Fanuc TP program (LS listing): POLIR.LS

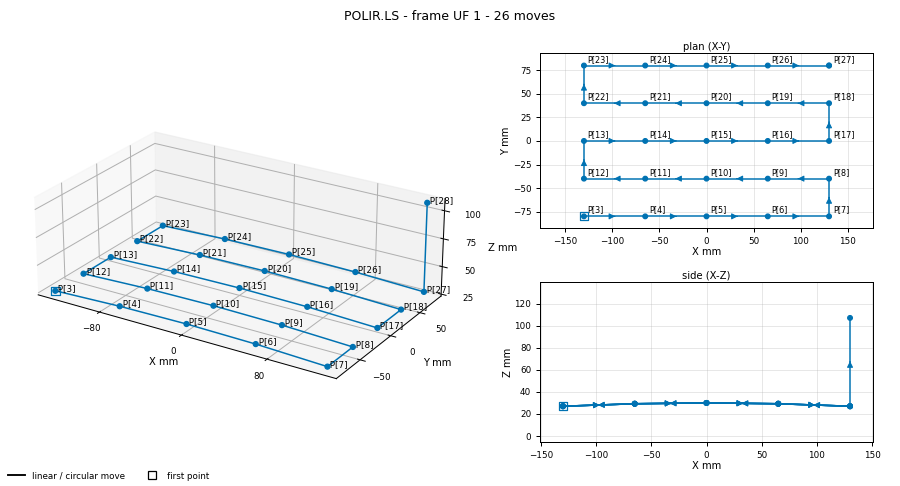
[picture p0: tool path of POLIR.LS in frame UF 1, 26 of 29 moves have a stored position in this frame; points joined in program order, loops and branches not executed]
/PROG  POLIR
/ATTR
OWNER		= MNEDITOR;
COMMENT		= "RoboDK sequence";
PROG_SIZE	= 0;
CREATE		= DATE 31-12-14  TIME 12:00:00;
MODIFIED	= DATE 31-12-14  TIME 12:00:00;
FILE_NAME	= POLIR;
VERSION		= 0;
LINE_COUNT	= 38;
MEMORY_SIZE	= 0;
PROTECT		= READ_WRITE;
TCD:  STACK_SIZE	= 0,
      TASK_PRIORITY	= 50,
      TIME_SLICE	= 0,
      BUSY_LAMP_OFF	= 0,
      ABORT_REQUEST	= 0,
      PAUSE_REQUEST	= 0;
DEFAULT_GROUP	= 1,*,*,*,*,*,*;
CONTROL_CODE	= 00000000 00000000;
/MN
   1:  ! Program generated by RoboDK v6.0.6 for FANUC M-10iD/12 on 24/ ;
   2:  ! 09/2026 00:37:20 ;
   3:  ! Using nominal kinematics. ;
   4:  UFRAME_NUM=1 ;
   5:  ! UF1:850.0,0.0,90.0,0.0,0.0,0.0 ;
   6:  UTOOL_NUM=1 ;
   7:  ! UT1:0.0,0.0,200.0,0.0,0.0,0.0 ;
   8:J P[1] 2% CNT1 ACC100 ;
   9:J P[2] 2% CNT1 ACC100 ;
  10:  DO[1]=ON ;
  11:L P[3] 40mm/sec CNT1 ACC100 ;
  12:L P[4] 40mm/sec CNT1 ACC100 ;
  13:L P[5] 40mm/sec CNT1 ACC100 ;
  14:L P[6] 40mm/sec CNT1 ACC100 ;
  15:L P[7] 40mm/sec CNT1 ACC100 ;
  16:L P[8] 40mm/sec CNT1 ACC100 ;
  17:L P[9] 40mm/sec CNT1 ACC100 ;
  18:L P[10] 40mm/sec CNT1 ACC100 ;
  19:L P[11] 40mm/sec CNT1 ACC100 ;
  20:L P[12] 40mm/sec CNT1 ACC100 ;
  21:L P[13] 40mm/sec CNT1 ACC100 ;
  22:L P[14] 40mm/sec CNT1 ACC100 ;
  23:L P[15] 40mm/sec CNT1 ACC100 ;
  24:L P[16] 40mm/sec CNT1 ACC100 ;
  25:L P[17] 40mm/sec CNT1 ACC100 ;
  26:L P[18] 40mm/sec CNT1 ACC100 ;
  27:L P[19] 40mm/sec CNT1 ACC100 ;
  28:L P[20] 40mm/sec CNT1 ACC100 ;
  29:L P[21] 40mm/sec CNT1 ACC100 ;
  30:L P[22] 40mm/sec CNT1 ACC100 ;
  31:L P[23] 40mm/sec CNT1 ACC100 ;
  32:L P[24] 40mm/sec CNT1 ACC100 ;
  33:L P[25] 40mm/sec CNT1 ACC100 ;
  34:L P[26] 40mm/sec CNT1 ACC100 ;
  35:L P[27] 40mm/sec CNT1 ACC100 ;
  36:L P[28] 40mm/sec CNT1 ACC100 ;
  37:  DO[1]=OFF ;
  38:J P[29] 2% CNT1 ACC100 ;
/POS
P[1]{
   GP1:
    UF : 1, UT : 1,
	J1=    -6.453 deg,	J2=    -8.040 deg,	J3=    -17.302 deg,
	J4=    -0.316 deg,	J5=    -70.069 deg,	J6=    6.554 deg
};
P[2]{
   GP1:
    UF : 1, UT : 1,
	J1=    -6.453 deg,	J2=    -6.370 deg,	J3=    -28.638 deg,
	J4=    -0.348 deg,	J5=    -58.733 deg,	J6=    6.627 deg
};
P[3]{
   GP1:
    UF : 1, UT : 1,        CONFIG : 'N U T, 0, 0, 0',
	X =  -130.000  mm,	Y =   -80.000  mm,	Z =    26.996  mm,
	W =   180.000 deg,	P =    -2.646 deg,	R =     0.000 deg
};
P[4]{
   GP1:
    UF : 1, UT : 1,        CONFIG : 'N U T, 0, 0, 0',
	X =   -65.000  mm,	Y =   -80.000  mm,	Z =    29.249  mm,
	W =   180.000 deg,	P =    -1.324 deg,	R =     0.000 deg
};
P[5]{
   GP1:
    UF : 1, UT : 1,        CONFIG : 'N U T, 0, 0, 0',
	X =     0.000  mm,	Y =   -80.000  mm,	Z =    30.000  mm,
	W =   180.000 deg,	P =     0.000 deg,	R =     0.000 deg
};
P[6]{
   GP1:
    UF : 1, UT : 1,        CONFIG : 'N U T, 0, 0, 0',
	X =    65.000  mm,	Y =   -80.000  mm,	Z =    29.249  mm,
	W =   180.000 deg,	P =     1.324 deg,	R =     0.000 deg
};
P[7]{
   GP1:
    UF : 1, UT : 1,        CONFIG : 'N U T, 0, 0, 0',
	X =   130.000  mm,	Y =   -80.000  mm,	Z =    26.996  mm,
	W =   180.000 deg,	P =     2.646 deg,	R =     0.000 deg
};
P[8]{
   GP1:
    UF : 1, UT : 1,        CONFIG : 'N U T, 0, 0, 0',
	X =   130.000  mm,	Y =   -40.000  mm,	Z =    26.996  mm,
	W =   180.000 deg,	P =     2.646 deg,	R =     0.000 deg
};
P[9]{
   GP1:
    UF : 1, UT : 1,        CONFIG : 'N U T, 0, 0, 0',
	X =    65.000  mm,	Y =   -40.000  mm,	Z =    29.249  mm,
	W =   180.000 deg,	P =     1.324 deg,	R =     0.000 deg
};
P[10]{
   GP1:
    UF : 1, UT : 1,        CONFIG : 'N U T, 0, 0, 0',
	X =     0.000  mm,	Y =   -40.000  mm,	Z =    30.000  mm,
	W =   180.000 deg,	P =     0.000 deg,	R =     0.000 deg
};
P[11]{
   GP1:
    UF : 1, UT : 1,        CONFIG : 'N U T, 0, 0, 0',
	X =   -65.000  mm,	Y =   -40.000  mm,	Z =    29.249  mm,
	W =   180.000 deg,	P =    -1.324 deg,	R =     0.000 deg
};
P[12]{
   GP1:
    UF : 1, UT : 1,        CONFIG : 'N U T, 0, 0, 0',
	X =  -130.000  mm,	Y =   -40.000  mm,	Z =    26.996  mm,
	W =   180.000 deg,	P =    -2.646 deg,	R =     0.000 deg
};
P[13]{
   GP1:
    UF : 1, UT : 1,        CONFIG : 'N U T, 0, 0, 0',
	X =  -130.000  mm,	Y =     0.000  mm,	Z =    26.996  mm,
	W =   180.000 deg,	P =    -2.646 deg,	R =     0.000 deg
};
P[14]{
   GP1:
    UF : 1, UT : 1,        CONFIG : 'N U T, 0, 0, 0',
	X =   -65.000  mm,	Y =     0.000  mm,	Z =    29.249  mm,
	W =   180.000 deg,	P =    -1.324 deg,	R =     0.000 deg
};
P[15]{
   GP1:
    UF : 1, UT : 1,        CONFIG : 'N U T, 0, 0, 0',
	X =     0.000  mm,	Y =     0.000  mm,	Z =    30.000  mm,
	W =   180.000 deg,	P =     0.000 deg,	R =     0.000 deg
};
P[16]{
   GP1:
    UF : 1, UT : 1,        CONFIG : 'N U T, 0, 0, 0',
	X =    65.000  mm,	Y =     0.000  mm,	Z =    29.249  mm,
	W =   180.000 deg,	P =     1.324 deg,	R =     0.000 deg
};
P[17]{
   GP1:
    UF : 1, UT : 1,        CONFIG : 'N U T, 0, 0, 0',
	X =   130.000  mm,	Y =     0.000  mm,	Z =    26.996  mm,
	W =   180.000 deg,	P =     2.646 deg,	R =     0.000 deg
};
P[18]{
   GP1:
    UF : 1, UT : 1,        CONFIG : 'N U T, 0, 0, 0',
	X =   130.000  mm,	Y =    40.000  mm,	Z =    26.996  mm,
	W =   180.000 deg,	P =     2.646 deg,	R =     0.000 deg
};
P[19]{
   GP1:
    UF : 1, UT : 1,        CONFIG : 'N U T, 0, 0, 0',
	X =    65.000  mm,	Y =    40.000  mm,	Z =    29.249  mm,
	W =   180.000 deg,	P =     1.324 deg,	R =     0.000 deg
};
P[20]{
   GP1:
    UF : 1, UT : 1,        CONFIG : 'N U T, 0, 0, 0',
	X =     0.000  mm,	Y =    40.000  mm,	Z =    30.000  mm,
	W =   180.000 deg,	P =     0.000 deg,	R =     0.000 deg
};
P[21]{
   GP1:
    UF : 1, UT : 1,        CONFIG : 'N U T, 0, 0, 0',
	X =   -65.000  mm,	Y =    40.000  mm,	Z =    29.249  mm,
	W =   180.000 deg,	P =    -1.324 deg,	R =     0.000 deg
};
P[22]{
   GP1:
    UF : 1, UT : 1,        CONFIG : 'N U T, 0, 0, 0',
	X =  -130.000  mm,	Y =    40.000  mm,	Z =    26.996  mm,
	W =   180.000 deg,	P =    -2.646 deg,	R =     0.000 deg
};
P[23]{
   GP1:
    UF : 1, UT : 1,        CONFIG : 'N U T, 0, 0, 0',
	X =  -130.000  mm,	Y =    80.000  mm,	Z =    26.996  mm,
	W =   180.000 deg,	P =    -2.646 deg,	R =     0.000 deg
};
P[24]{
   GP1:
    UF : 1, UT : 1,        CONFIG : 'N U T, 0, 0, 0',
	X =   -65.000  mm,	Y =    80.000  mm,	Z =    29.249  mm,
	W =   180.000 deg,	P =    -1.324 deg,	R =     0.000 deg
};
P[25]{
   GP1:
    UF : 1, UT : 1,        CONFIG : 'N U T, 0, 0, 0',
	X =     0.000  mm,	Y =    80.000  mm,	Z =    30.000  mm,
	W =   180.000 deg,	P =     0.000 deg,	R =     0.000 deg
};
P[26]{
   GP1:
    UF : 1, UT : 1,        CONFIG : 'N U T, 0, 0, 0',
	X =    65.000  mm,	Y =    80.000  mm,	Z =    29.249  mm,
	W =   180.000 deg,	P =     1.324 deg,	R =     0.000 deg
};
P[27]{
   GP1:
    UF : 1, UT : 1,        CONFIG : 'N U T, 0, 0, 0',
	X =   130.000  mm,	Y =    80.000  mm,	Z =    26.996  mm,
	W =   180.000 deg,	P =     2.646 deg,	R =     0.000 deg
};
P[28]{
   GP1:
    UF : 1, UT : 1,        CONFIG : 'N U T, 0, 0, 0',
	X =   130.000  mm,	Y =    80.000  mm,	Z =   106.996  mm,
	W =   180.000 deg,	P =     2.646 deg,	R =     0.000 deg
};
P[29]{
   GP1:
    UF : 1, UT : 1,
	J1=    -6.453 deg,	J2=    -8.040 deg,	J3=    -17.302 deg,
	J4=    -0.316 deg,	J5=    -70.069 deg,	J6=    6.554 deg
};
/END
